// TIA Portal V19 export
VAR_GLOBAL   // PLC tag table "Safety"
   DI_Door_1_Lock AT %I12.0 : Bool;
   DI_Door_2_Lock AT %I12.1 : Bool;
   DI_Door_3_Lock AT %I12.2 : Bool;
   DI_Door_4_Lock AT %I12.3 : Bool;
   DI_Door_5_Lock AT %I12.4 : Bool;
   DI_Door_6_Lock AT %I12.5 : Bool;
   DI_Door_7_Lock AT %I12.6 : Bool;
   DI_Door_8_Lock AT %I12.7 : Bool;
   DQ_Door_1_Lock AT %Q16.0 : Bool;
   DQ_Door_2_Lock AT %Q16.1 : Bool;
   DQ_Door_3_Lock AT %Q16.2 : Bool;
   DQ_Door_4_Lock AT %Q16.3 : Bool;
   DQ_Door_5_Lock AT %Q16.4 : Bool;
   DQ_Door_6_Lock AT %Q16.5 : Bool;
   DQ_Door_7_Lock AT %Q16.6 : Bool;
   DQ_Door_8_Lock AT %Q16.7 : Bool;
END_VAR
